(* IEC 61131-3 sources: sis-interlock-demo/src/DUTs/Generated, 1 file *)

(* ---- ST_SisIo.dut.st ---- *)
// AUTO-GENERATED by cemgen 1.0.0 — не редактировать: правьте матрицу и запустите
//   python -m cemgen generate <файл матрицы .csv или .xlsx>
// Матрица: SIS-V101-CEM, объект V-101, ревизия B от 2026-10-19, SHA-256 сетки df2ed4841a9453ca
// Назначение: образ ввода-вывода ПАЗ объекта V-101: токи датчиков 4–20 мА, дискретные входы с
//             контролем линии, ключи и кнопка, выходы-разрешения xQ* (TRUE — под напряжением).
//             Поля — по тегам матрицы (DESIGN.md, 9.3), порядок — первое появление каналов, затем
//             ключи и выходы.
// Автор:      kr0nsch; код — генератор cemgen
// Версия:     1.0.0
// Документ:   docs/DESIGN.md, раздел «10. Генератор cemgen»; docs/cause_effect_matrix.md
// ВНИМАНИЕ:   код демонстрационный и не предназначен для систем безопасности. Реальная ПАЗ требует
//             определения SIL, сертифицированных аппаратных и программных средств и валидации по
//             ГОСТ Р МЭК 61511.
{attribute 'qualified_only'}
TYPE ST_SisIo :
STRUCT
    // --- 1 PSHH101: Давление в V-101 аварийно высокое (ai, 2oo3) ---
    rPT101A_mA : REAL;   // PT101A, мА: шкала 0…1,6 МПа; 1 PSHH101, 2 PSLL101
    rPT101B_mA : REAL;   // PT101B, мА: шкала 0…1,6 МПа; 1 PSHH101, 2 PSLL101
    rPT101C_mA : REAL;   // PT101C, мА: шкала 0…1,6 МПа; 1 PSHH101, 2 PSLL101
    // --- 3 LSHH102: Уровень жидкости в V-101 аварийно высокий (ai, 2oo3) ---
    rLT102A_mA : REAL;   // LT102A, мА: шкала 0…2,4 м; 3 LSHH102, 4 LSLL102
    rLT102B_mA : REAL;   // LT102B, мА: шкала 0…2,4 м; 3 LSHH102, 4 LSLL102
    rLT102C_mA : REAL;   // LT102C, мА: шкала 0…2,4 м; 3 LSHH102, 4 LSLL102
    // --- 5 TSHH103: Температура жидкости в V-101 аварийно высокая (ai, 1oo2) ---
    rTT103A_mA : REAL;   // TT103A, мА: шкала 0…150 °C; 5 TSHH103
    rTT103B_mA : REAL;   // TT103B, мА: шкала 0…150 °C; 5 TSHH103
    // --- 6 ASHH104: Загазованность у V-101 аварийно высокая (ai, 2oo3) ---
    rAT104A_mA : REAL;   // AT104A, мА: шкала 0…100 % НКПР; 6 ASHH104
    rAT104B_mA : REAL;   // AT104B, мА: шкала 0…100 % НКПР; 6 ASHH104
    rAT104C_mA : REAL;   // AT104C, мА: шкала 0…100 % НКПР; 6 ASHH104
    // --- 7 BSH105: Пожар у V-101 (di, 1oo2) ---
    xBS105A    : BOOL;   // BS105A: норма 1; 7 BSH105
    xBS105A_Ok : BOOL;   // BS105A: контроль линии, TRUE — исправна
    xBS105B    : BOOL;   // BS105B: норма 1; 7 BSH105
    xBS105B_Ok : BOOL;   // BS105B: контроль линии, TRUE — исправна
    // --- 8 HS106: Аварийный останов кнопкой (di, 1oo2) ---
    xHS106A    : BOOL;   // HS106A: норма 1; 8 HS106
    xHS106A_Ok : BOOL;   // HS106A: контроль линии, TRUE — исправна
    xHS106B    : BOOL;   // HS106B: норма 1; 8 HS106
    xHS106B_Ok : BOOL;   // HS106B: контроль линии, TRUE — исправна
    // --- 9 PSLL108: Давление воздуха КИП аварийно низкое (di, 2oo2) ---
    xPS108A    : BOOL;   // PS108A: норма 1; 9 PSLL108
    xPS108A_Ok : BOOL;   // PS108A: контроль линии, TRUE — исправна
    xPS108B    : BOOL;   // PS108B: норма 1; 9 PSLL108
    xPS108B_Ok : BOOL;   // PS108B: контроль линии, TRUE — исправна
    // --- 10 ESL109: Потеря напряжения щита 0,4 кВ (di, 1oo1) ---
    xES109     : BOOL;   // ES109: норма 1; 10 ESL109
    xES109_Ok  : BOOL;   // ES109: контроль линии, TRUE — исправна
    // --- ключи и кнопка ---
    xHS120     : BOOL;   // HS120: кнопка «Сброс ПАЗ» (действует фронт)
    xHS121     : BOOL;   // HS121: ключ «Разрешение байпасов»
    xHS122     : BOOL;   // HS122: ключ «Разрешение пусковых обходов»
    // --- выходы ПАЗ: разрешения, обесточивание на срабатывание ---
    xQESDV101  : BOOL;   // ESDV101: разрешение, TRUE — под напряжением; FALSE — закрыт
    xQBDV101   : BOOL;   // BDV101: разрешение, TRUE — под напряжением; FALSE — открыт
    xQESDV102  : BOOL;   // ESDV102: разрешение, TRUE — под напряжением; FALSE — закрыт
    xQP101A    : BOOL;   // P101A: разрешение, TRUE — под напряжением; FALSE — остановлен
    xQP101B    : BOOL;   // P101B: разрешение, TRUE — под напряжением; FALSE — остановлен
    xQH101     : BOOL;   // H101: разрешение, TRUE — под напряжением; FALSE — отключён
    xQUA110    : BOOL;   // UA110: разрешение, TRUE — под напряжением; FALSE — сигнал
END_STRUCT
END_TYPE
